// TIA Portal V20 export
TYPE "Afag_ist_Werte"
   STRUCT
      Telegram_identifier : Byte;
      operating_mode : Byte;   // manufacturer-specific
      PROFIDRIVE_Statusword : Word;
      actual_position : DInt;   // transmitted parameters in default-parameterization
      actual_speed : DInt;   // transmitted parameters in default-parameterization
      active_current_actual_value : DInt;   // transmitted parameters in default-parameterization
      digital_Inputs : DInt;   // transmitted parameters in default-parameterization
   END_STRUCT;
END_TYPE
